{region 'Documentation'}
(*!
<summary>Check that IN is strictly earlier than Maximum.</summary>
<description>

A value at or beyond 24 hours reports Error before comparison or baseline capture.

</description>
*)
{endregion}
FUNCTION_BLOCK AssertEarlierThan_LTOD EXTENDS AssertionBase
VAR_INPUT
    IN : LTOD; //! Actual value checked or observed by this Assertion.
    Maximum : LTOD; //! Exclusive upper bound; the actual value or count must be smaller.
END_VAR

SUPER^();

{region 'Documentation'}
(*!
<summary>Evaluate the typed temporal relation and report higher-priority errors first.</summary>
*)
{endregion}
METHOD PROTECTED Assert
VAR
    Message : STRING(GVL_Constants.MessageLength);
    MaximumText : STRING(GVL_Constants.AssertionValueLength);
    ActualText : STRING(GVL_Constants.AssertionValueLength);
END_VAR
IF NOT EvaluationActive THEN
    RETURN;
END_IF;

IF Result = E_Result.Error THEN
    RETURN;
END_IF;

IF NOT IsTimeOfDayValid_LTOD(Value := IN) THEN
    Error(Message := 'Assertion error: IN is outside the valid LTOD range (less than 24 hours).');
    RETURN;
END_IF;

IF NOT IsTimeOfDayValid_LTOD(Value := Maximum) THEN
    Error(Message := 'Assertion error: Maximum is outside the valid LTOD range (less than 24 hours).');
    RETURN;
END_IF;

IF Result = E_Result.Failed THEN
    RETURN;
END_IF;

IF IN >= Maximum THEN
    MaximumText := LTOD_TO_STRING(Maximum);
    ActualText := LTOD_TO_STRING(IN);
    Message := CONCAT('Assertion failed: value is not earlier than limit. Maximum = ',
        MaximumText);
    Message := CONCAT(Message, ', Actual = ');
    Message := CONCAT(Message, ActualText);
    Message := CONCAT(Message, '.');
    Fail(Message := Message);
    RETURN;
END_IF;

Pass();
END_METHOD

END_FUNCTION_BLOCK

(* stored: Version 1.1.0.1
   POU AssertEarlierThan_LTOD: Id {3784ff6e-3e89-44ed-8bf8-2813298ab11d}, SpecialFunc None
   Folder Internal: Id {683a2f71-b44e-4aa1-ae92-8a0a331d03a8}
   Method Assert: Id {150668b6-e3e7-4a8b-9c95-4fbe378939d3} *)
